(* IEC 61131-3 sources: llm-plc-st-eval/data/definitivo/qwen2.5-coder_14b/B3/zero_shot, 3 files *)

(* ---- ejec_1.st ---- *)
```pascal
FUNCTION_BLOCK FB_Contador
VAR_INPUT
    sensorPieza : BOOL; // Sensor fotoeléctrico que detecta la pieza
    btnReset : BOOL;    // Botón de reset para reiniciar el contador
END_VAR

VAR_OUTPUT
    loteListo : BOOL; // Salida que indica que se ha completado un lote
    cuenta : INT;      // Contador de piezas
END_VAR

VAR
    sensorAnterior : BOOL; // Variable para almacenar el estado anterior del sensor
END_VAR

// Inicialización del sensorAnterior con el valor actual del sensorPieza
IF sensorPieza THEN
    sensorAnterior := TRUE;
ELSE
    sensorAnterior := FALSE;
END_IF

// Lógica de conteo
IF sensorPieza AND NOT sensorAnterior THEN
    cuenta := cuenta + 1;
END_IF

// Actualización del sensorAnterior
sensorAnterior := sensorPieza;

// Lógica para detectar el lote completo
IF cuenta >= 12 THEN
    loteListo := TRUE;
ELSE
    loteListo := FALSE;
END_IF

// Lógica de reset
IF btnReset THEN
    cuenta := 0;
    loteListo := FALSE;
END_IF
END_FUNCTION_BLOCK
```

(* ---- ejec_2.st ---- *)
```pascal
FUNCTION_BLOCK FB_Contador
VAR_INPUT
    sensorPieza : BOOL; // Entrada del sensor fotoeléctrico
    btnReset : BOOL; // Botón de reset
END_VAR

VAR_OUTPUT
    loteListo : BOOL; // Salida de lote completo
    cuenta : INT; // Contador de piezas
END_VAR

VAR
    sensorAnterior : BOOL; // Estado anterior del sensor
END_VAR

// Inicialización
IF sensorAnterior = FALSE AND sensorPieza = TRUE THEN
    cuenta := cuenta + 1; // Incrementar el contador
END_IF;

// Reset
IF btnReset THEN
    cuenta := 0; // Poner el contador en cero
    loteListo := FALSE; // Desactivar la salida de lote
END_IF;

// Control de lote completo
IF cuenta >= 12 THEN
    loteListo := TRUE; // Activar la salida de lote completo
ELSE
    loteListo := FALSE; // Desactivar la salida de lote completo
END_IF;

// Actualizar el estado anterior del sensor
sensorAnterior := sensorPieza;
```

Este código implementa un FUNCTION_BLOCK que cuenta piezas en una línea de producción según las especificaciones proporcionadas. Utiliza una variable interna `sensorAnterior` para detectar transiciones del sensor fotoeléctrico. El contador se incrementa cada vez que se detecta una pieza, y se resetea cuando se presiona el botón de reset. La salida de lote completo se activa cuando se alcanzan 12 piezas.

(* ---- ejec_3.st ---- *)
```pascal
FUNCTION_BLOCK FB_Contador
VAR_INPUT
    sensorPieza : BOOL; // Sensor fotoeléctrico que detecta la pieza
    btnReset : BOOL;    // Botón de reset para reiniciar el contador
END_VAR

VAR_OUTPUT
    loteListo : BOOL;  // Salida que indica que se ha completado un lote
    cuenta : INT;       // Contador de piezas
END_VAR

VAR
    sensorAnterior : BOOL; // Variable para almacenar el estado anterior del sensor
END_VAR

// Inicialización de variables
IF sensorAnterior = FALSE AND sensorPieza = TRUE THEN
    cuenta := cuenta + 1; // Incrementar el contador al detectar una pieza
END_IF;

// Control del botón de reset
IF btnReset THEN
    cuenta := 0; // Reiniciar el contador
    loteListo := FALSE; // Desactivar la salida de lote completo
END_IF;

// Control de la salida de lote completo
IF cuenta >= 12 THEN
    loteListo := TRUE; // Activar la salida de lote completo
ELSE
    loteListo := FALSE; // Desactivar la salida de lote completo si no se han completado 12 piezas
END_IF;

// Actualizar el estado anterior del sensor
sensorAnterior := sensorPieza;
END_FUNCTION_BLOCK
```
